(* IEC 61131-3 sources: sis-interlock-demo/tests/GVLs, 2 files *)

(* ---- GVL_TestsSis.gvl.st ---- *)
// Назначение: экземпляры наборов тестов логики ПАЗ, написанных вручную (граничные случаи, раздел
//             12.3). Объявление экземпляра регистрирует набор в coUnit; PRG_Tests их не перечисляет.
//             {attribute 'linkalways'} обязателен: на GVL никто не ссылается, и без атрибута CODESYS
//             3.5.17 не включает её в приложение — наборы молча не выполняются.
// Автор:      kr0nsch
// Версия:     0.1.0
// Документ:   docs/DESIGN.md, раздел «12.3 Граничные случаи (вручную, команда A)»
// ВНИМАНИЕ:   код демонстрационный и не предназначен для систем безопасности. Реальная ПАЗ
//             требует определения SIL, сертифицированных аппаратных и программных средств
//             и валидации по ГОСТ Р МЭК 61511.
{attribute 'qualified_only'}
{attribute 'linkalways'}
VAR_GLOBAL
    fbVoteEvalTest    : FB_VoteEval_Test;      // F_VoteEval, F_VoteArchChannels, F_VoteArchRequired
    fbVotingTest      : FB_Voting_Test;        // FB_Voting, F_VoteCheckCfg
    fbCauseEffectTest : FB_CauseEffect_Test;   // FB_CauseEffect, F_CemCheckCfg
    fbSisEventLogTest : FB_SisEventLog_Test;   // FB_SisEventLog, I_SisEventSink
    fbSisUnitTest     : FB_SisUnit_Test;       // FB_SisUnit
    fbSisUtilTest     : FB_SisUtil_Test;       // CRC, биты, NE 43, масштабирование, F_SisLogEvent
    fbCommonTest      : FB_Common_Test;        // пределы, умолчания, коды перечислений, размеры
END_VAR

(* ---- GVL_TestsTruthTables.gvl.st ---- *)
// AUTO-GENERATED by tools_project/gen_voting_tests.py — не редактировать: правьте генератор или модель
//   tools_project/vote_model.py и запустите python tools_project/gen_voting_tests.py
// Назначение: экземпляры сгенерированных наборов таблиц истинности голосования. Объявление
//             экземпляра регистрирует набор в coUnit; {attribute 'linkalways'} обязателен: на GVL
//             никто не ссылается, без атрибута CODESYS 3.5.17 не включает её в приложение.
// Автор:      kr0nsch; код — генератор tools_project/gen_voting_tests.py
// Версия:     0.1.0
// Документ:   docs/DESIGN.md, раздел «12.2 Таблицы истинности (генерируются)»
// ВНИМАНИЕ:   код демонстрационный и не предназначен для систем безопасности. Реальная ПАЗ
//             требует определения SIL, сертифицированных аппаратных и программных средств
//             и валидации по ГОСТ Р МЭК 61511.
{attribute 'qualified_only'}
{attribute 'linkalways'}
VAR_GLOBAL
    fbVoteTableEvalTest     : FB_VoteTableEval_Test;       // F_VoteEval: 12 таблиц, 300 строк
    fbVoteTable2oo3VTDITest : FB_VoteTable2oo3VTDI_Test;   // FB_Voting: 2oo3 VT DI, 512 строк
    fbVoteTable2oo3VTAITest : FB_VoteTable2oo3VTAI_Test;   // FB_Voting: 2oo3 VT AI, 512 строк
    fbVoteTable2oo3DSDITest : FB_VoteTable2oo3DSDI_Test;   // FB_Voting: 2oo3 DS DI, 512 строк
    fbVoteTable2oo3DSAITest : FB_VoteTable2oo3DSAI_Test;   // FB_Voting: 2oo3 DS AI, 512 строк
    fbVoteTable2oo3DADITest : FB_VoteTable2oo3DADI_Test;   // FB_Voting: 2oo3 DA DI, 512 строк
    fbVoteTable2oo3DAAITest : FB_VoteTable2oo3DAAI_Test;   // FB_Voting: 2oo3 DA AI, 512 строк
    fbVoteTableFbSmallTest  : FB_VoteTableFbSmall_Test;    // FB_Voting: 1oo1, 1oo2, 2oo2
END_VAR
